TYPE ST_HallInputs :
STRUCT
    bUpperButton : BOOL;
    bLowerButton : BOOL;
END_STRUCT
END_TYPE

(* stored: Version 1.1.0.1
   DUT ST_HallInputs: Id {90a41573-756d-42f1-9774-06324dce6a31} *)
